Staubli VAL3: teachHome.pgx

public program teachHome()
  local bool l_bResult
begin
  l_bResult=userPageConfirm("是否记录当前位置为home位置？")
  if l_bResult
    savedata:jHome=herej()
    savedata:libSave()
    delay(0.1)
    popUpMsg("home位置已记录并保存")
  endIf
end
